Fanuc KAREL source: kt00474.KL

-- PROVISIONAL review KL for V1013-1; original PC SHA256 048b88de654025c002eceb735755ccb025ce42fb74608fa853c81e43c3362846
-- Incomplete behavior may be omitted. Consult companion uncertainty JSON. Do not deploy.
PROGRAM KT00474
%NOLOCKGROUP
-- UNRESOLVED_DECL P1 type=000101
-- UNRESOLVED_DECL P2 type=000101
-- UNRESOLVED_DECL OUT type=000101
BEGIN
  -- UNRESOLVED_PC offsets 5-29; opcodes 49,49,60,4A
  -- UNRESOLVED_PC offsets 34-38; opcodes 7F
END KT00474
